SUBAPPLICATION Input_Toggle_RPC_TO_Remote_AX_OPC (* Wie Input_Toggle_RPC_TO_Remote_QXA_OPC, aber ohne logiBUS_QXA: der Zustand geht als AX-Plug STATE nach aussen *)
  (* Standard: 61499-2; Description: Copyright (c) 2026 Meisterschulen am Ostbahnhof This program and the accompanying materials are made available under the terms of the Eclipse Public License 2.0 which is available at https://www.eclipse.org/legal/epl-2.0/ SPDX-License-Identifier: EPL-2.0 *)
  (* Version 1.0, 2026-10-18, Franz Höpfinger, Meisterschulen am Ostbahnhof, Ohne QXA: AX_SUBSCRIBE_1.OUT direkt auf den Plug STATE, Anzeige/Weiterverarbeitung frei waehlbar *)
  PACKAGE MyLib::sys;
  IMPORT logiBUS::io::DI::logiBUS_DI;
  IMPORT logiBUS::io::DI::logiBUS_DI_S;
  IMPORT logiBUS::io::DI::logiBUS_DI_Events::BUTTON_PRESS_DOWN;
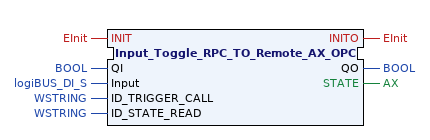
  EVENT_INPUT
    INIT : EInit; (* Initialization Request *)
  END_EVENT
  EVENT_OUTPUT
    INITO : EInit; (* Initialization Confirm *)
  END_EVENT
  VAR_INPUT
    QI : BOOL := TRUE; (* Quality Input - TRUE to enable service *)
    Input : logiBUS::io::DI::logiBUS_DI_S := logiBUS_DI::Invalid; (* Taster Input_I1..I8 (Tastendruck ruft die Methode) *)
    ID_TRIGGER_CALL : WSTRING; (* Methodenadresse (ACTION=CALL_METHOD, mit Endpunkt) *)
    ID_STATE_READ : WSTRING; (* Lokale Adresse (BOOL, ACTION=READ) fuer den Zustand *)
  END_VAR
  VAR_OUTPUT
    QO : BOOL; (* Quality Output - TRUE if service executed successfully *)
  END_VAR
  PLUGS
    STATE : adapter::types::unidirectional::AX; (* Flipflop-Zustand (lokal gelesen) *)
  END_PLUGS
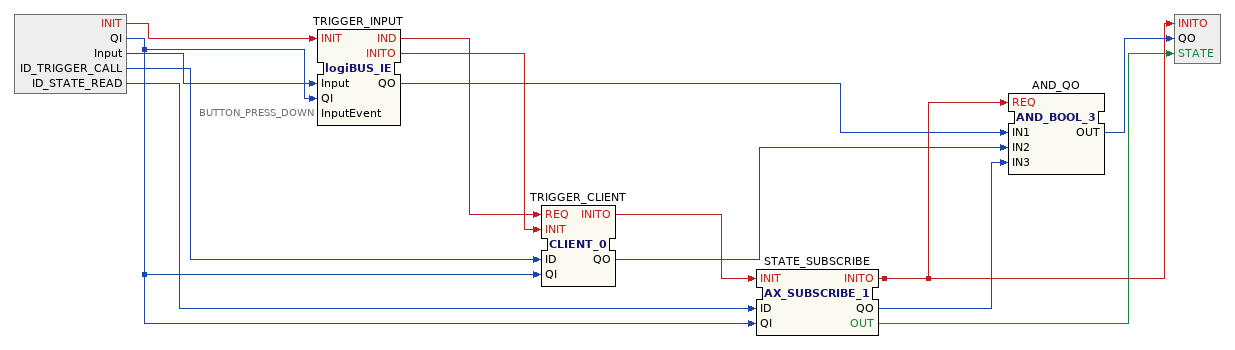
  FBS
    TRIGGER_INPUT : logiBUS::io::DI::logiBUS_IE(InputEvent := BUTTON_PRESS_DOWN);
    TRIGGER_CLIENT : iec61499::net::CLIENT_0;
    STATE_SUBSCRIBE : adapter::net::AX_SUBSCRIBE_1;
    AND_QO : iec61131::booleanOperators::AND_BOOL_3;
  END_FBS
  EVENT_CONNECTIONS
    TRIGGER_INPUT.IND TO TRIGGER_CLIENT.REQ;
    INIT TO TRIGGER_INPUT.INIT;
    TRIGGER_INPUT.INITO TO TRIGGER_CLIENT.INIT;
    TRIGGER_CLIENT.INITO TO STATE_SUBSCRIBE.INIT;
    STATE_SUBSCRIBE.INITO TO INITO;
    STATE_SUBSCRIBE.INITO TO AND_QO.REQ;
  END_CONNECTIONS
  DATA_CONNECTIONS
    Input TO TRIGGER_INPUT.Input;
    ID_TRIGGER_CALL TO TRIGGER_CLIENT.ID;
    ID_STATE_READ TO STATE_SUBSCRIBE.ID;
    QI TO TRIGGER_INPUT.QI;
    QI TO TRIGGER_CLIENT.QI;
    QI TO STATE_SUBSCRIBE.QI;
    TRIGGER_INPUT.QO TO AND_QO.IN1;
    TRIGGER_CLIENT.QO TO AND_QO.IN2;
    STATE_SUBSCRIBE.QO TO AND_QO.IN3;
    AND_QO.OUT TO QO;
  END_CONNECTIONS
  ADAPTER_CONNECTIONS
    STATE_SUBSCRIBE.OUT TO STATE;
  END_CONNECTIONS
END_SUBAPPLICATION
